(* IEC 61131-3 sources: llm-plc-st-eval/data/definitivo/qwen2.5-coder_14b/A3/zero_shot, 3 files *)

(* ---- ejec_1.st ---- *)
```pascal
FUNCTION_BLOCK FB_Com
VAR_INPUT
    txReq : BOOL;  // Petición de transmisión
    rxOk  : BOOL;  // Confirmación de recepción correcta
    rxData: INT;   // Datos recibidos
END_VAR

VAR_OUTPUT
    txData : INT;  // Datos a transmitir
    ocupado: BOOL;  // Indica si el sistema está ocupado
    ok     : BOOL;  // Indica si el intercambio fue exitoso
    error  : BOOL;  // Indica si el intercambio falló
    nIntentos: INT; // Número de intentos realizados
END_VAR

VAR
    estado    : INT := 0; // Estado actual del intercambio
    intentos  : INT := 0; // Contador de intentos
    timer     : TON;      // Temporizador para el plazo de 500 ms
    valorTx   : INT := 0; // Valor a transmitir
    inicioInt : BOOL := FALSE; // Indica si se ha iniciado un intento
END_VAR

// Estado 0: Esperando petición de transmisión
IF txReq AND NOT inicioInt THEN
    estado := 1;
    intentos := 1;
    nIntentos := intentos;
    valorTx := 100;
    txData := valorTx;
    ocupado := TRUE;
    ok := FALSE;
    error := FALSE;
    timer(IN := TRUE, PT := T#500MS);
    inicioInt := TRUE;
END_IF

// Estado 1: Esperando respuesta
IF estado = 1 THEN
    IF rxOk AND rxData = valorTx THEN
        estado := 2;
        ok := TRUE;
        ocupado := FALSE;
    ELSIF timer.Q THEN
        IF intentos < 3 THEN
            intentos := intentos + 1;
            nIntentos := intentos;
            timer(IN := TRUE, PT := T#500MS);
        ELSE
            estado := 3;
            error := TRUE;
            ocupado := FALSE;
        END_IF
    END_IF
END_IF

// Estado 2: Intercambio exitoso
IF estado = 2 THEN
    // Mantener ok activo hasta la siguiente petición
END_IF

// Estado 3: Intercambio fallido
IF estado = 3 THEN
    // Mantener error activo hasta la siguiente petición
END_IF

// Reiniciar el estado si se recibe una nueva petición mientras se está ocupado
IF txReq AND inicioInt THEN
    // Ignorar la nueva petición
END_IF

// Reiniciar el estado al finalizar el intercambio
IF estado = 2 OR estado = 3 THEN
    inicioInt := FALSE;
END_IF
END_FUNCTION_BLOCK
```

(* ---- ejec_2.st ---- *)
```pascal
FUNCTION_BLOCK FB_Com
VAR_INPUT
    txReq : BOOL;  // Petición de transmisión
    rxOk  : BOOL;  // Confirmación de recepción
    rxData: INT;   // Datos recibidos
END_VAR

VAR_OUTPUT
    txData  : INT;  // Datos a transmitir
    ocupado : BOOL; // Estado de ocupado
    ok      : BOOL; // Estado de éxito
    error   : BOOL; // Estado de error
    nIntentos: INT; // Número de intentos
END_VAR

VAR
    estado    : INT := 0; // Estado actual del intercambio
    intentos  : INT := 0; // Contador de intentos
    tiempoEspera: TON; // Temporizador para el plazo de espera
    valorTx   : INT := 0; // Valor a transmitir
END_VAR

// Inicialización del temporizador
tiempoEspera(IN := FALSE, PT := T#500MS);

// Máquina de estados
CASE estado OF
    0: // Estado inicial
        IF txReq THEN
            valorTx := 100; // Valor de prueba
            txData := valorTx;
            ocupado := TRUE;
            intentos := 1;
            nIntentos := intentos;
            tiempoEspera(IN := TRUE); // Iniciar temporizador
            estado := 1; // Pasar al estado de espera de respuesta
        END_IF

    1: // Estado de espera de respuesta
        IF rxOk AND (rxData = valorTx) THEN
            ok := TRUE;
            ocupado := FALSE;
            estado := 0; // Terminar intercambio
        ELSIF tiempoEspera.Q THEN
            IF intentos < 3 THEN
                intentos := intentos + 1;
                nIntentos := intentos;
                tiempoEspera(IN := TRUE); // Reiniciar temporizador
            ELSE
                error := TRUE;
                ocupado := FALSE;
                estado := 0; // Terminar intercambio
            END_IF
        END_IF

    ELSE
        estado := 0; // Restablecer estado en caso de error
END_CASE

// Mantener ok y error activos hasta el siguiente intercambio
IF estado = 0 THEN
    ok := FALSE;
    error := FALSE;
END_IF
```

Este código implementa una máquina de estados para manejar el intercambio de petición/respuesta con un dispositivo externo, siguiendo los requisitos especificados.

(* ---- ejec_3.st ---- *)
```pascal
FUNCTION_BLOCK FB_Com
VAR_INPUT
    txReq : BOOL;  // Petición de transmisión
    rxOk  : BOOL;  // Confirmación de recepción
    rxData: INT;   // Datos recibidos
END_VAR

VAR_OUTPUT
    txData  : INT;  // Datos a transmitir
    ocupado : BOOL; // Indica si se está ocupado en un intercambio
    ok      : BOOL; // Indica si el intercambio fue exitoso
    error   : BOOL; // Indica si el intercambio falló
    nIntentos: INT;  // Número de intentos realizados
END_VAR

VAR
    estado    : INT := 0; // Estado del intercambio (0: Idle, 1: Enviando, 2: Esperando respuesta)
    intentos  : INT := 0; // Contador de intentos
    timer     : TON;     // Temporizador para esperar la respuesta
    valorTx   : INT := 0; // Valor a transmitir
    inicioIntercambio : BOOL := FALSE; // Indica si se ha iniciado un intercambio
END_VAR

// Inicialización del temporizador
timer(IN := FALSE, PT := T#500MS);

// Máquina de estados
CASE estado OF
    0: // Estado Idle
        IF txReq AND NOT inicioIntercambio THEN
            inicioIntercambio := TRUE;
            estado := 1;
            intentos := 1;
            nIntentos := intentos;
            valorTx := 100;
            txData := valorTx;
            ocupado := TRUE;
            timer(IN := TRUE);
        END_IF

    1: // Estado Enviando
        IF rxOk AND (rxData = valorTx) THEN
            estado := 0;
            ok := TRUE;
            ocupado := FALSE;
            inicioIntercambio := FALSE;
        ELSIF timer.Q THEN
            IF intentos < 3 THEN
                intentos := intentos + 1;
                nIntentos := intentos;
                timer(IN := TRUE);
            ELSE
                estado := 0;
                error := TRUE;
                ocupado := FALSE;
                inicioIntercambio := FALSE;
            END_IF
        END_IF

    2: // Estado Esperando respuesta
        // Este estado no se utiliza en este código, pero se mantiene por claridad.
        // El estado de espera se maneja en el estado 1.
END_CASE

// Mantener ok y error activos hasta el siguiente intercambio
IF estado = 0 THEN
    IF ok THEN
        ok := FALSE;
    END_IF
    IF error THEN
        error := FALSE;
    END_IF
END_IF
```
